(* IEC 61131-3 sources: plc-iiot-stack/src/POUs/Iiot/F_IiotQuality, 2 files *)

(* ---- F_IiotQuality.decl.st ---- *)
// Назначение: качество метрики по статусу NE 107 и достоверности устройства (data_schema 3.2):
//             F — bad; S, C — uncertain; Good, M — good при достоверном значении, иначе bad.
// Автор:      kr0nsch
// Версия:     0.1.0
// Документ:   docs/plc_mqtt.md, раздел «Телеметрия»
FUNCTION F_IiotQuality : E_IiotQuality
VAR_INPUT
    xValid : BOOL;   // значение достоверно (выход xValid AI и DI; для двигателя — TRUE)
    iNe107 : INT;    // код E_Ne107Status устройства (0 Good ... 4 Failure)
END_VAR

(* ---- F_IiotQuality.impl.st ---- *)
IF iNe107 >= TO_INT(E_IiotNe107.Failure) THEN
    F_IiotQuality := E_IiotQuality.Bad;
ELSIF iNe107 = TO_INT(E_IiotNe107.OutOfSpecification) OR iNe107 = TO_INT(E_IiotNe107.CheckFunction) THEN
    F_IiotQuality := E_IiotQuality.Uncertain;
ELSIF xValid THEN
    F_IiotQuality := E_IiotQuality.Good;
ELSE
    F_IiotQuality := E_IiotQuality.Bad;
END_IF
